Universal Robots URScript: T006_codellama_34b_adversarial_A8.6_rep1.urscript

def bin_picking():
    # Home position
    movej(p[0, 0, -90, 0, 180, 0], a=350.0, v=400.0)

    # Above bin
    movel(p[-200, 0, 0, 0, 0, 0], a=350.0, v=400.0)

    # Descend
